(* IEC 61131-3 sources: tsplc/packages/vscode-extension/tests/fixtures/blueprint/transport/FB_ZoneConveyor, 1 file *)

(* ---- FB_ZoneConveyor.declaration.st ---- *)
FUNCTION_BLOCK FB_ZoneConveyor
VAR_IN_OUT
	Conveyor : ST_Conveyor;
END_VAR
VAR
	pConveyor : POINTER TO ST_Conveyor;
END_VAR
